(* IEC 61131-3 sources: kns-port-domestic/tools/plcopen/tests/fixtures/constructs/src/POUs/F_Sum, 2 files *)

(* ---- F_Sum.decl.st ---- *)
// Назначение: сумма элементов массива любой длины (VAR_IN_OUT CONSTANT, ARRAY[*])
// Автор:      <ИМЯ ФАМИЛИЯ>
// Версия:     0.1.0
// Документ:   docs/plcopen.md
FUNCTION F_Sum : LREAL
VAR_IN_OUT CONSTANT
    arValues : ARRAY[*] OF REAL;
END_VAR
VAR
    diIdx : DINT;
END_VAR

(* ---- F_Sum.impl.st ---- *)
F_Sum := 0;
FOR diIdx := LOWER_BOUND(arValues, 1) TO UPPER_BOUND(arValues, 1) DO
    F_Sum := F_Sum + arValues[diIdx];
END_FOR
